{attribute 'qualified_only'}
{attribute 'strict'}
{attribute 'to_string'}
TYPE E_AxisControlCommand : (
    None := 0,
    MoveAbsolute := 1,
    MoveRelative := 2,
    Jog := 3,
    Home := 4,
    Stop := 5,
    SetAbsolutePosition := 6
);
END_TYPE

(* stored: Version 1.1.0.1, ProductVersion 3.1.4026.20
   DUT E_AxisControlCommand: Id {2d4682f8-7f06-5d45-bef6-1af034a59ec2} *)
